Fanuc KAREL source: IO0193.KL

PROGRAM IO0193
%NOLOCKGROUP
%ENVIRONMENT REGOPE
ROUTINE RTEST
VAR
  I : INTEGER
  STATUS : INTEGER
  ENTRY : INTEGER
  A : ARRAY[3] OF INTEGER
  B : BOOLEAN
  R : REAL
  P : XYZWPR
  JPOS : JOINTPOS
  PF : POSITION
BEGIN
  I = 1
  A[1] = 2
  B = TRUE
  R = 1.0
  P = GET_POS_REG(1,STATUS,1)
END RTEST
BEGIN
  RTEST
END IO0193
